FUNCTION_BLOCK FB_SafeEStop
VAR_INPUT
END_VAR
VAR_OUTPUT
	bSafeState:		BOOL;
	bIsReset:		BOOL;
	fbError:		FB_Error;
END_VAR
VAR
	{attribute 'displaymode':='binary'}
	nDiag	AT %I*:	UINT;
	nState	AT %I*:	USINT;
	sMsg:			STRING;
	i:				INT;
END_VAR

bSafeState := nState = 3;
bIsReset := nState = 5;
CASE nState OF
	0: //undefined
		IF NOT fbError.bError THEN
			fbError.M_Set(1, 'Undefinierter State!', nState, eID := E_ErrorIDs.eUndefinedState, eSrc := E_ErrorSrcs.eSafetyFb);
		END_IF
	1: //RUN
		IF fbError.bError THEN
			fbError.M_Reset();
		END_IF
	2:;
	3:;
	4://Error
		IF NOT fbError.bError THEN
			IF nDiag.0 THEN
				sMsg := CONCAT(sMsg, 'DiskrepGr1,');
			END_IF
			IF nDiag.1 THEN
				sMsg := CONCAT(sMsg, 'DiskrepGr2,');
			END_IF
			IF nDiag.2 THEN
				sMsg := CONCAT(sMsg, 'DiskrepGrSec,');
			END_IF
			IF nDiag.4 THEN
				sMsg := CONCAT(sMsg, 'EDM1,');
			END_IF
			IF nDiag.5 THEN
				sMsg := CONCAT(sMsg, 'EDM2,');
			END_IF
			IF nDiag.8 THEN
				sMsg := CONCAT(sMsg, 'DiskrepErrGr1Plus');
			END_IF
			IF nDiag.9 THEN
				sMsg := CONCAT(sMsg, 'DiskrepErrGr2Plus');
			END_IF
			IF nDiag.10 THEN
				sMsg := CONCAT(sMsg, 'DiskrepErrSecPlus');
			END_IF
			
			fbError.M_Set(1, sMsg, TO_INT(nDiag), eID := E_ErrorIDs.eSafetyFbError, eSrc := E_ErrorSrcs.eSafetyFb);
		END_IF
	5,6,7,8,9:;
	ELSE //undefined
		IF NOT fbError.bError THEN
			fbError.M_Set(1, 'Undefinierter State!', nState, eID := E_ErrorIDs.eUndefinedState, eSrc := E_ErrorSrcs.eSafetyFb);
		END_IF
END_CASE

END_FUNCTION_BLOCK

(* stored: Version 1.1.0.1, ProductVersion 3.1.4024.9
   POU FB_SafeEStop: Id {68d26bd3-3af4-4021-a28c-8acef07f86f3}, SpecialFunc None *)
